(* IEC 61131-3 sources: kns-port-domestic/upstream/kns-pump-station/src/GVLs/Generated, 7 files *)

(* ---- GVL_CfgProject.gvl.st ---- *)
// AUTO-GENERATED by iolistgen 0.2.0 — не редактировать; источник: 03_io_list.csv
// SHA-256 перечня 06336d13c4b2; генератор st-codesys
// Назначение: уставки проекта — Cfg устройств из перечня сигналов, те же инициализаторы, что у GVL_Persist.
// PRG_ApplyProjectCfg копирует их в GVL_Persist (контракт plc-process-lib 18.3, правило 2).
{attribute 'qualified_only'}
VAR_GLOBAL CONSTANT
    // --- dev_no 11: P101 — Насос Н1 (MotorVfd) ---
    // lint:allow STL007 структура-константа: имя как у GVL_Persist.stP101Cfg (контракт 18.3, правило 2)
    stP101Cfg : PL.ST_MotorCfg := (
        tFbStart := T#10S,
        tFbStop := T#15S,
        tMinStop := T#30S,
        uiMaxStartsPerHour := 10,
        stVfd := (
            rSpeedMin_pct := 60.0,
            rRampUp_pctps := 5.0,
            rRampDown_pctps := 5.0,
            xFbFromComm := FALSE,
            xCommLossIsFault := FALSE
        ),
        udiAlarmIdBase := 110
    );
    // --- dev_no 12: P102 — Насос Н2 (MotorVfd) ---
    // lint:allow STL007 структура-константа: имя как у GVL_Persist.stP102Cfg (контракт 18.3, правило 2)
    stP102Cfg : PL.ST_MotorCfg := (
        tFbStart := T#10S,
        tFbStop := T#15S,
        tMinStop := T#30S,
        uiMaxStartsPerHour := 10,
        stVfd := (
            rSpeedMin_pct := 60.0,
            rRampUp_pctps := 5.0,
            rRampDown_pctps := 5.0,
            xFbFromComm := FALSE,
            xCommLossIsFault := FALSE
        ),
        udiAlarmIdBase := 120
    );
    // --- dev_no 13: P103 — Насос Н3 (MotorVfd) ---
    // lint:allow STL007 структура-константа: имя как у GVL_Persist.stP103Cfg (контракт 18.3, правило 2)
    stP103Cfg : PL.ST_MotorCfg := (
        tFbStart := T#10S,
        tFbStop := T#15S,
        tMinStop := T#30S,
        uiMaxStartsPerHour := 10,
        stVfd := (
            rSpeedMin_pct := 60.0,
            rRampUp_pctps := 5.0,
            rRampDown_pctps := 5.0,
            xFbFromComm := FALSE,
            xCommLossIsFault := FALSE
        ),
        udiAlarmIdBase := 130
    );
    // --- dev_no 14: V1 — Вытяжной вентилятор В1 павильона (Motor) ---
    // lint:allow STL007 структура-константа: имя как у GVL_Persist.stV1Cfg (контракт 18.3, правило 2)
    stV1Cfg : PL.ST_MotorCfg := (
        tMinStop := T#10S,
        udiAlarmIdBase := 140,
        astAlarm := [
            (ePriority := PL.E_AlarmPriority.Low),  // 0 FailToStart
            (ePriority := PL.E_AlarmPriority.Low),  // 1 FeedbackLost
            (ePriority := PL.E_AlarmPriority.High),  // 2 FailToStop
            (ePriority := PL.E_AlarmPriority.High),  // 3 UncommandedRun
            (ePriority := PL.E_AlarmPriority.Low),  // 4 ExtFault
            (ePriority := PL.E_AlarmPriority.None),  // 5 InterlockTrip
            (ePriority := PL.E_AlarmPriority.Medium),  // 6 CommLoss
            (ePriority := PL.E_AlarmPriority.Low)  // 7 SpeedDeviation
        ]
    );
    // --- dev_no 101: LT101 — Уровень в приёмном резервуаре (AnalogInput) ---
    // lint:allow STL007 структура-константа: имя как у GVL_Persist.stLT101Cfg (контракт 18.3, правило 2)
    stLT101Cfg : PL.ST_AnalogInputCfg := (
        rRangeHi_eu := 5.0,
        tFilter := T#2S,
        astLimit := [
            (xEnable := TRUE, rSetpoint_eu := 4.0, rHyst_eu := 0.05, tOnDelay := T#3S),  // 0 HH
            (xEnable := TRUE, rSetpoint_eu := 3.5, rHyst_eu := 0.05, tOnDelay := T#3S),  // 1 H
            (xEnable := TRUE, rSetpoint_eu := 0.8, rHyst_eu := 0.05, tOnDelay := T#3S),  // 2 L
            (xEnable := TRUE, rSetpoint_eu := 0.5, rHyst_eu := 0.05, tOnDelay := T#3S)  // 3 LL
        ],
        udiAlarmIdBase := 1010,
        astAlarm := [
            (ePriority := PL.E_AlarmPriority.High),  // 0 HH
            (ePriority := PL.E_AlarmPriority.Medium),  // 1 H
            (ePriority := PL.E_AlarmPriority.Medium),  // 2 L
            (ePriority := PL.E_AlarmPriority.High),  // 3 LL
            (ePriority := PL.E_AlarmPriority.Medium),  // 4 Failure
            (ePriority := PL.E_AlarmPriority.Low),  // 5 OutOfRange
            (ePriority := PL.E_AlarmPriority.None),  // 6 (резерв)
            (ePriority := PL.E_AlarmPriority.None)  // 7 (резерв)
        ]
    );
    // --- dev_no 102: LS102 — Поплавок «аварийно высокий уровень» (H, 4,2 м) (DigitalInput) ---
    // lint:allow STL007 структура-константа: имя как у GVL_Persist.stLS102Cfg (контракт 18.3, правило 2)
    stLS102Cfg : PL.ST_DigitalInputCfg := (
        xInvert := TRUE,
        tOnDelay := T#2S,
        udiAlarmIdBase := 1020,
        astAlarm := [
            (ePriority := PL.E_AlarmPriority.High),  // 0 State
            (ePriority := PL.E_AlarmPriority.Medium),  // 1 Failure
            (ePriority := PL.E_AlarmPriority.None),  // 2 (резерв)
            (ePriority := PL.E_AlarmPriority.None),  // 3 (резерв)
            (ePriority := PL.E_AlarmPriority.None),  // 4 (резерв)
            (ePriority := PL.E_AlarmPriority.None),  // 5 (резерв)
            (ePriority := PL.E_AlarmPriority.None),  // 6 (резерв)
            (ePriority := PL.E_AlarmPriority.None)  // 7 (резерв)
        ]
    );
    // --- dev_no 103: LS103 — Поплавок «сухой ход» (L, 0,4 м) (DigitalInput) ---
    // lint:allow STL007 структура-константа: имя как у GVL_Persist.stLS103Cfg (контракт 18.3, правило 2)
    stLS103Cfg : PL.ST_DigitalInputCfg := (
        xInvert := TRUE,
        tOnDelay := T#1S,
        eFailValue := PL.E_DiFailValue.ForceTrue,
        udiAlarmIdBase := 1030,
        astAlarm := [
            (ePriority := PL.E_AlarmPriority.High),  // 0 State
            (ePriority := PL.E_AlarmPriority.Medium),  // 1 Failure
            (ePriority := PL.E_AlarmPriority.None),  // 2 (резерв)
            (ePriority := PL.E_AlarmPriority.None),  // 3 (резерв)
            (ePriority := PL.E_AlarmPriority.None),  // 4 (резерв)
            (ePriority := PL.E_AlarmPriority.None),  // 5 (резерв)
            (ePriority := PL.E_AlarmPriority.None),  // 6 (резерв)
            (ePriority := PL.E_AlarmPriority.None)  // 7 (резерв)
        ]
    );
    // --- dev_no 111: IT111 — Насос Н1: ток двигателя (измеряет ПЧ) (AnalogInput) ---
    // lint:allow STL007 структура-константа: имя как у GVL_Persist.stIT111Cfg (контракт 18.3, правило 2)
    stIT111Cfg : PL.ST_AnalogInputCfg := (
        eInput := PL.E_AiInputType.Raw,
        rRangeHi_eu := 60.0,
        rRawHi_cnt := 600.0,
        tFilter := T#1S,
        astLimit := [
            (xEnable := TRUE, rSetpoint_eu := 34.0, tOnDelay := T#10S),  // 0 HH
            (xEnable := TRUE, rSetpoint_eu := 31.0, tOnDelay := T#10S),  // 1 H
            (xEnable := FALSE),  // 2 L
            (xEnable := FALSE)  // 3 LL
        ],
        udiAlarmIdBase := 1110,
        astAlarm := [
            (ePriority := PL.E_AlarmPriority.Medium),  // 0 HH
            (ePriority := PL.E_AlarmPriority.Low),  // 1 H
            (ePriority := PL.E_AlarmPriority.Low),  // 2 L
            (ePriority := PL.E_AlarmPriority.Medium),  // 3 LL
            (ePriority := PL.E_AlarmPriority.Medium),  // 4 Failure
            (ePriority := PL.E_AlarmPriority.Low),  // 5 OutOfRange
            (ePriority := PL.E_AlarmPriority.None),  // 6 (резерв)
            (ePriority := PL.E_AlarmPriority.None)  // 7 (резерв)
        ]
    );
    // --- dev_no 112: TS112 — Насос Н1: перегрев обмотки (термовыключатели, реле защиты насоса) (DigitalInput) ---
    // lint:allow STL007 структура-константа: имя как у GVL_Persist.stTS112Cfg (контракт 18.3, правило 2)
    stTS112Cfg : PL.ST_DigitalInputCfg := (
        xInvert := TRUE,
        udiAlarmIdBase := 1120,
        astAlarm := [
            (ePriority := PL.E_AlarmPriority.High),  // 0 State
            (ePriority := PL.E_AlarmPriority.Medium),  // 1 Failure
            (ePriority := PL.E_AlarmPriority.None),  // 2 (резерв)
            (ePriority := PL.E_AlarmPriority.None),  // 3 (резерв)
            (ePriority := PL.E_AlarmPriority.None),  // 4 (резерв)
            (ePriority := PL.E_AlarmPriority.None),  // 5 (резерв)
            (ePriority := PL.E_AlarmPriority.None),  // 6 (резерв)
            (ePriority := PL.E_AlarmPriority.None)  // 7 (резерв)
        ]
    );
    // --- dev_no 113: MS113 — Насос Н1: протечка в камеру статора (датчик влажности, реле защиты на… (DigitalInput) ---
    // lint:allow STL007 структура-константа: имя как у GVL_Persist.stMS113Cfg (контракт 18.3, правило 2)
    stMS113Cfg : PL.ST_DigitalInputCfg := (
        tOnDelay := T#10S,
        udiAlarmIdBase := 1130,
        astAlarm := [
            (ePriority := PL.E_AlarmPriority.Medium),  // 0 State
            (ePriority := PL.E_AlarmPriority.Medium),  // 1 Failure
            (ePriority := PL.E_AlarmPriority.None),  // 2 (резерв)
            (ePriority := PL.E_AlarmPriority.None),  // 3 (резерв)
            (ePriority := PL.E_AlarmPriority.None),  // 4 (резерв)
            (ePriority := PL.E_AlarmPriority.None),  // 5 (резерв)
            (ePriority := PL.E_AlarmPriority.None),  // 6 (резерв)
            (ePriority := PL.E_AlarmPriority.None)  // 7 (резерв)
        ]
    );
    // --- dev_no 121: IT121 — Насос Н2: ток двигателя (измеряет ПЧ) (AnalogInput) ---
    // lint:allow STL007 структура-константа: имя как у GVL_Persist.stIT121Cfg (контракт 18.3, правило 2)
    stIT121Cfg : PL.ST_AnalogInputCfg := (
        eInput := PL.E_AiInputType.Raw,
        rRangeHi_eu := 60.0,
        rRawHi_cnt := 600.0,
        tFilter := T#1S,
        astLimit := [
            (xEnable := TRUE, rSetpoint_eu := 34.0, tOnDelay := T#10S),  // 0 HH
            (xEnable := TRUE, rSetpoint_eu := 31.0, tOnDelay := T#10S),  // 1 H
            (xEnable := FALSE),  // 2 L
            (xEnable := FALSE)  // 3 LL
        ],
        udiAlarmIdBase := 1210,
        astAlarm := [
            (ePriority := PL.E_AlarmPriority.Medium),  // 0 HH
            (ePriority := PL.E_AlarmPriority.Low),  // 1 H
            (ePriority := PL.E_AlarmPriority.Low),  // 2 L
            (ePriority := PL.E_AlarmPriority.Medium),  // 3 LL
            (ePriority := PL.E_AlarmPriority.Medium),  // 4 Failure
            (ePriority := PL.E_AlarmPriority.Low),  // 5 OutOfRange
            (ePriority := PL.E_AlarmPriority.None),  // 6 (резерв)
            (ePriority := PL.E_AlarmPriority.None)  // 7 (резерв)
        ]
    );
    // --- dev_no 122: TS122 — Насос Н2: перегрев обмотки (термовыключатели, реле защиты насоса) (DigitalInput) ---
    // lint:allow STL007 структура-константа: имя как у GVL_Persist.stTS122Cfg (контракт 18.3, правило 2)
    stTS122Cfg : PL.ST_DigitalInputCfg := (
        xInvert := TRUE,
        udiAlarmIdBase := 1220,
        astAlarm := [
            (ePriority := PL.E_AlarmPriority.High),  // 0 State
            (ePriority := PL.E_AlarmPriority.Medium),  // 1 Failure
            (ePriority := PL.E_AlarmPriority.None),  // 2 (резерв)
            (ePriority := PL.E_AlarmPriority.None),  // 3 (резерв)
            (ePriority := PL.E_AlarmPriority.None),  // 4 (резерв)
            (ePriority := PL.E_AlarmPriority.None),  // 5 (резерв)
            (ePriority := PL.E_AlarmPriority.None),  // 6 (резерв)
            (ePriority := PL.E_AlarmPriority.None)  // 7 (резерв)
        ]
    );
    // --- dev_no 123: MS123 — Насос Н2: протечка в камеру статора (датчик влажности, реле защиты на… (DigitalInput) ---
    // lint:allow STL007 структура-константа: имя как у GVL_Persist.stMS123Cfg (контракт 18.3, правило 2)
    stMS123Cfg : PL.ST_DigitalInputCfg := (
        tOnDelay := T#10S,
        udiAlarmIdBase := 1230,
        astAlarm := [
            (ePriority := PL.E_AlarmPriority.Medium),  // 0 State
            (ePriority := PL.E_AlarmPriority.Medium),  // 1 Failure
            (ePriority := PL.E_AlarmPriority.None),  // 2 (резерв)
            (ePriority := PL.E_AlarmPriority.None),  // 3 (резерв)
            (ePriority := PL.E_AlarmPriority.None),  // 4 (резерв)
            (ePriority := PL.E_AlarmPriority.None),  // 5 (резерв)
            (ePriority := PL.E_AlarmPriority.None),  // 6 (резерв)
            (ePriority := PL.E_AlarmPriority.None)  // 7 (резерв)
        ]
    );
    // --- dev_no 131: IT131 — Насос Н3: ток двигателя (измеряет ПЧ) (AnalogInput) ---
    // lint:allow STL007 структура-константа: имя как у GVL_Persist.stIT131Cfg (контракт 18.3, правило 2)
    stIT131Cfg : PL.ST_AnalogInputCfg := (
        eInput := PL.E_AiInputType.Raw,
        rRangeHi_eu := 60.0,
        rRawHi_cnt := 600.0,
        tFilter := T#1S,
        astLimit := [
            (xEnable := TRUE, rSetpoint_eu := 34.0, tOnDelay := T#10S),  // 0 HH
            (xEnable := TRUE, rSetpoint_eu := 31.0, tOnDelay := T#10S),  // 1 H
            (xEnable := FALSE),  // 2 L
            (xEnable := FALSE)  // 3 LL
        ],
        udiAlarmIdBase := 1310,
        astAlarm := [
            (ePriority := PL.E_AlarmPriority.Medium),  // 0 HH
            (ePriority := PL.E_AlarmPriority.Low),  // 1 H
            (ePriority := PL.E_AlarmPriority.Low),  // 2 L
            (ePriority := PL.E_AlarmPriority.Medium),  // 3 LL
            (ePriority := PL.E_AlarmPriority.Medium),  // 4 Failure
            (ePriority := PL.E_AlarmPriority.Low),  // 5 OutOfRange
            (ePriority := PL.E_AlarmPriority.None),  // 6 (резерв)
            (ePriority := PL.E_AlarmPriority.None)  // 7 (резерв)
        ]
    );
    // --- dev_no 132: TS132 — Насос Н3: перегрев обмотки (термовыключатели, реле защиты насоса) (DigitalInput) ---
    // lint:allow STL007 структура-константа: имя как у GVL_Persist.stTS132Cfg (контракт 18.3, правило 2)
    stTS132Cfg : PL.ST_DigitalInputCfg := (
        xInvert := TRUE,
        udiAlarmIdBase := 1320,
        astAlarm := [
            (ePriority := PL.E_AlarmPriority.High),  // 0 State
            (ePriority := PL.E_AlarmPriority.Medium),  // 1 Failure
            (ePriority := PL.E_AlarmPriority.None),  // 2 (резерв)
            (ePriority := PL.E_AlarmPriority.None),  // 3 (резерв)
            (ePriority := PL.E_AlarmPriority.None),  // 4 (резерв)
            (ePriority := PL.E_AlarmPriority.None),  // 5 (резерв)
            (ePriority := PL.E_AlarmPriority.None),  // 6 (резерв)
            (ePriority := PL.E_AlarmPriority.None)  // 7 (резерв)
        ]
    );
    // --- dev_no 133: MS133 — Насос Н3: протечка в камеру статора (датчик влажности, реле защиты на… (DigitalInput) ---
    // lint:allow STL007 структура-константа: имя как у GVL_Persist.stMS133Cfg (контракт 18.3, правило 2)
    stMS133Cfg : PL.ST_DigitalInputCfg := (
        tOnDelay := T#10S,
        udiAlarmIdBase := 1330,
        astAlarm := [
            (ePriority := PL.E_AlarmPriority.Medium),  // 0 State
            (ePriority := PL.E_AlarmPriority.Medium),  // 1 Failure
            (ePriority := PL.E_AlarmPriority.None),  // 2 (резерв)
            (ePriority := PL.E_AlarmPriority.None),  // 3 (резерв)
            (ePriority := PL.E_AlarmPriority.None),  // 4 (резерв)
            (ePriority := PL.E_AlarmPriority.None),  // 5 (резерв)
            (ePriority := PL.E_AlarmPriority.None),  // 6 (резерв)
            (ePriority := PL.E_AlarmPriority.None)  // 7 (резерв)
        ]
    );
    // --- dev_no 201: PT201 — Давление в напорном коллекторе (AnalogInput) ---
    // lint:allow STL007 структура-константа: имя как у GVL_Persist.stPT201Cfg (контракт 18.3, правило 2)
    stPT201Cfg : PL.ST_AnalogInputCfg := (
        rRangeHi_eu := 10.0,
        tFilter := T#1S,
        astLimit := [
            (xEnable := TRUE, rSetpoint_eu := 5.0, tOnDelay := T#5S),  // 0 HH
            (xEnable := TRUE, rSetpoint_eu := 4.0, tOnDelay := T#5S),  // 1 H
            (xEnable := TRUE, rSetpoint_eu := 1.0, rHyst_eu := 0.1, tOnDelay := T#5S),  // 2 L
            (xEnable := TRUE, rSetpoint_eu := 0.5, rHyst_eu := 0.1, tOnDelay := T#5S)  // 3 LL
        ],
        udiAlarmIdBase := 2010,
        astAlarm := [
            (ePriority := PL.E_AlarmPriority.High),  // 0 HH
            (ePriority := PL.E_AlarmPriority.Medium),  // 1 H
            (ePriority := PL.E_AlarmPriority.Medium),  // 2 L
            (ePriority := PL.E_AlarmPriority.High),  // 3 LL
            (ePriority := PL.E_AlarmPriority.Medium),  // 4 Failure
            (ePriority := PL.E_AlarmPriority.Low),  // 5 OutOfRange
            (ePriority := PL.E_AlarmPriority.None),  // 6 (резерв)
            (ePriority := PL.E_AlarmPriority.None)  // 7 (резерв)
        ]
    );
    // --- dev_no 202: FT202 — Расход в напорном коллекторе (AnalogInput) ---
    // lint:allow STL007 структура-константа: имя как у GVL_Persist.stFT202Cfg (контракт 18.3, правило 2)
    stFT202Cfg : PL.ST_AnalogInputCfg := (
        rRangeHi_eu := 500.0,
        rLowCut_pct := 1.0,
        tFilter := T#3S,
        astLimit := [
            (xEnable := FALSE),  // 0 HH
            (xEnable := FALSE),  // 1 H
            (xEnable := TRUE, rSetpoint_eu := 30.0, rHyst_eu := 5.0, tOnDelay := T#30S),  // 2 L
            (xEnable := FALSE)  // 3 LL
        ],
        udiAlarmIdBase := 2020,
        astAlarm := [
            (ePriority := PL.E_AlarmPriority.High),  // 0 HH
            (ePriority := PL.E_AlarmPriority.Low),  // 1 H
            (ePriority := PL.E_AlarmPriority.Medium),  // 2 L
            (ePriority := PL.E_AlarmPriority.High),  // 3 LL
            (ePriority := PL.E_AlarmPriority.Medium),  // 4 Failure
            (ePriority := PL.E_AlarmPriority.Low),  // 5 OutOfRange
            (ePriority := PL.E_AlarmPriority.None),  // 6 (резерв)
            (ePriority := PL.E_AlarmPriority.None)  // 7 (резерв)
        ]
    );
    // --- dev_no 203: LS203 — Затопление камеры задвижек (DigitalInput) ---
    // lint:allow STL007 структура-константа: имя как у GVL_Persist.stLS203Cfg (контракт 18.3, правило 2)
    stLS203Cfg : PL.ST_DigitalInputCfg := (
        tOnDelay := T#5S,
        udiAlarmIdBase := 2030,
        astAlarm := [
            (ePriority := PL.E_AlarmPriority.Medium),  // 0 State
            (ePriority := PL.E_AlarmPriority.Medium),  // 1 Failure
            (ePriority := PL.E_AlarmPriority.None),  // 2 (резерв)
            (ePriority := PL.E_AlarmPriority.None),  // 3 (резерв)
            (ePriority := PL.E_AlarmPriority.None),  // 4 (резерв)
            (ePriority := PL.E_AlarmPriority.None),  // 5 (резерв)
            (ePriority := PL.E_AlarmPriority.None),  // 6 (резерв)
            (ePriority := PL.E_AlarmPriority.None)  // 7 (резерв)
        ]
    );
    // --- dev_no 301: ES301 — Напряжение на вводе в норме (реле контроля фаз) (DigitalInput) ---
    // lint:allow STL007 структура-константа: имя как у GVL_Persist.stES301Cfg (контракт 18.3, правило 2)
    stES301Cfg : PL.ST_DigitalInputCfg := (
        tOnDelay := T#3S,
        xAlarmOnTrue := FALSE,
        udiAlarmIdBase := 3010,
        astAlarm := [
            (ePriority := PL.E_AlarmPriority.High),  // 0 State
            (ePriority := PL.E_AlarmPriority.Medium),  // 1 Failure
            (ePriority := PL.E_AlarmPriority.None),  // 2 (резерв)
            (ePriority := PL.E_AlarmPriority.None),  // 3 (резерв)
            (ePriority := PL.E_AlarmPriority.None),  // 4 (резерв)
            (ePriority := PL.E_AlarmPriority.None),  // 5 (резерв)
            (ePriority := PL.E_AlarmPriority.None),  // 6 (резерв)
            (ePriority := PL.E_AlarmPriority.None)  // 7 (резерв)
        ]
    );
    // --- dev_no 302: YS302 — ИБП шкафа управления: работа от батарей (DigitalInput) ---
    // lint:allow STL007 структура-константа: имя как у GVL_Persist.stYS302Cfg (контракт 18.3, правило 2)
    stYS302Cfg : PL.ST_DigitalInputCfg := (
        tOnDelay := T#5S,
        udiAlarmIdBase := 3020,
        astAlarm := [
            (ePriority := PL.E_AlarmPriority.Medium),  // 0 State
            (ePriority := PL.E_AlarmPriority.Medium),  // 1 Failure
            (ePriority := PL.E_AlarmPriority.None),  // 2 (резерв)
            (ePriority := PL.E_AlarmPriority.None),  // 3 (резерв)
            (ePriority := PL.E_AlarmPriority.None),  // 4 (резерв)
            (ePriority := PL.E_AlarmPriority.None),  // 5 (резерв)
            (ePriority := PL.E_AlarmPriority.None),  // 6 (резерв)
            (ePriority := PL.E_AlarmPriority.None)  // 7 (резерв)
        ]
    );
    // --- dev_no 303: YS303 — ИБП шкафа управления: неисправность или разряд батарей (DigitalInput) ---
    // lint:allow STL007 структура-константа: имя как у GVL_Persist.stYS303Cfg (контракт 18.3, правило 2)
    stYS303Cfg : PL.ST_DigitalInputCfg := (
        tOnDelay := T#5S,
        udiAlarmIdBase := 3030,
        astAlarm := [
            (ePriority := PL.E_AlarmPriority.Medium),  // 0 State
            (ePriority := PL.E_AlarmPriority.Medium),  // 1 Failure
            (ePriority := PL.E_AlarmPriority.None),  // 2 (резерв)
            (ePriority := PL.E_AlarmPriority.None),  // 3 (резерв)
            (ePriority := PL.E_AlarmPriority.None),  // 4 (резерв)
            (ePriority := PL.E_AlarmPriority.None),  // 5 (резерв)
            (ePriority := PL.E_AlarmPriority.None),  // 6 (резерв)
            (ePriority := PL.E_AlarmPriority.None)  // 7 (резерв)
        ]
    );
    // --- dev_no 401: AT401 — Концентрация сероводорода H₂S в павильоне (AnalogInput) ---
    // lint:allow STL007 структура-константа: имя как у GVL_Persist.stAT401Cfg (контракт 18.3, правило 2)
    stAT401Cfg : PL.ST_AnalogInputCfg := (
        rRangeHi_eu := 40.0,
        astLimit := [
            (xEnable := TRUE, rSetpoint_eu := 10.0, rHyst_eu := 0.5, tOnDelay := T#5S),  // 0 HH
            (xEnable := TRUE, rSetpoint_eu := 5.0, rHyst_eu := 0.5, tOnDelay := T#5S),  // 1 H
            (xEnable := FALSE),  // 2 L
            (xEnable := FALSE)  // 3 LL
        ],
        udiAlarmIdBase := 4010,
        astAlarm := [
            (ePriority := PL.E_AlarmPriority.High),  // 0 HH
            (ePriority := PL.E_AlarmPriority.Medium),  // 1 H
            (ePriority := PL.E_AlarmPriority.Medium),  // 2 L
            (ePriority := PL.E_AlarmPriority.High),  // 3 LL
            (ePriority := PL.E_AlarmPriority.Medium),  // 4 Failure
            (ePriority := PL.E_AlarmPriority.Low),  // 5 OutOfRange
            (ePriority := PL.E_AlarmPriority.None),  // 6 (резерв)
            (ePriority := PL.E_AlarmPriority.None)  // 7 (резерв)
        ]
    );
    // --- dev_no 402: AT402 — Концентрация метана CH₄ в павильоне (AnalogInput) ---
    // lint:allow STL007 структура-константа: имя как у GVL_Persist.stAT402Cfg (контракт 18.3, правило 2)
    stAT402Cfg : PL.ST_AnalogInputCfg := (
        astLimit := [
            (xEnable := TRUE, rSetpoint_eu := 20.0, rHyst_eu := 1.0, tOnDelay := T#5S),  // 0 HH
            (xEnable := TRUE, rSetpoint_eu := 10.0, rHyst_eu := 1.0, tOnDelay := T#5S),  // 1 H
            (xEnable := FALSE),  // 2 L
            (xEnable := FALSE)  // 3 LL
        ],
        udiAlarmIdBase := 4020,
        astAlarm := [
            (ePriority := PL.E_AlarmPriority.High),  // 0 HH
            (ePriority := PL.E_AlarmPriority.Medium),  // 1 H
            (ePriority := PL.E_AlarmPriority.Medium),  // 2 L
            (ePriority := PL.E_AlarmPriority.High),  // 3 LL
            (ePriority := PL.E_AlarmPriority.Medium),  // 4 Failure
            (ePriority := PL.E_AlarmPriority.Low),  // 5 OutOfRange
            (ePriority := PL.E_AlarmPriority.None),  // 6 (резерв)
            (ePriority := PL.E_AlarmPriority.None)  // 7 (резерв)
        ]
    );
    // --- dev_no 403: TT403 — Температура воздуха в павильоне (AnalogInput) ---
    // lint:allow STL007 структура-константа: имя как у GVL_Persist.stTT403Cfg (контракт 18.3, правило 2)
    stTT403Cfg : PL.ST_AnalogInputCfg := (
        eInput := PL.E_AiInputType.Eng,
        rRangeLo_eu := -40.0,
        rRangeHi_eu := 60.0,
        astLimit := [
            (xEnable := FALSE),  // 0 HH
            (xEnable := TRUE, rSetpoint_eu := 35.0, rHyst_eu := 1.0, tOnDelay := T#1M),  // 1 H
            (xEnable := TRUE, rSetpoint_eu := 5.0, rHyst_eu := 1.0, tOnDelay := T#1M),  // 2 L
            (xEnable := FALSE)  // 3 LL
        ],
        udiAlarmIdBase := 4030,
        astAlarm := [
            (ePriority := PL.E_AlarmPriority.Low),  // 0 HH
            (ePriority := PL.E_AlarmPriority.Low),  // 1 H
            (ePriority := PL.E_AlarmPriority.Low),  // 2 L
            (ePriority := PL.E_AlarmPriority.Low),  // 3 LL
            (ePriority := PL.E_AlarmPriority.Medium),  // 4 Failure
            (ePriority := PL.E_AlarmPriority.Low),  // 5 OutOfRange
            (ePriority := PL.E_AlarmPriority.None),  // 6 (резерв)
            (ePriority := PL.E_AlarmPriority.None)  // 7 (резерв)
        ]
    );
    // --- dev_no 404: ZS404 — Дверь павильона открыта (DigitalInput) ---
    // lint:allow STL007 структура-константа: имя как у GVL_Persist.stZS404Cfg (контракт 18.3, правило 2)
    stZS404Cfg : PL.ST_DigitalInputCfg := (
        tOnDelay := T#2S,
        udiAlarmIdBase := 4040,
        astAlarm := [
            (ePriority := PL.E_AlarmPriority.Low),  // 0 State
            (ePriority := PL.E_AlarmPriority.Medium),  // 1 Failure
            (ePriority := PL.E_AlarmPriority.None),  // 2 (резерв)
            (ePriority := PL.E_AlarmPriority.None),  // 3 (резерв)
            (ePriority := PL.E_AlarmPriority.None),  // 4 (резерв)
            (ePriority := PL.E_AlarmPriority.None),  // 5 (резерв)
            (ePriority := PL.E_AlarmPriority.None),  // 6 (резерв)
            (ePriority := PL.E_AlarmPriority.None)  // 7 (резерв)
        ]
    );
    // --- dev_no 405: YS405 — Пожар (сигнал прибора пожарной сигнализации) (DigitalInput) ---
    // lint:allow STL007 структура-константа: имя как у GVL_Persist.stYS405Cfg (контракт 18.3, правило 2)
    stYS405Cfg : PL.ST_DigitalInputCfg := (
        udiAlarmIdBase := 4050,
        astAlarm := [
            (ePriority := PL.E_AlarmPriority.High),  // 0 State
            (ePriority := PL.E_AlarmPriority.Medium),  // 1 Failure
            (ePriority := PL.E_AlarmPriority.None),  // 2 (резерв)
            (ePriority := PL.E_AlarmPriority.None),  // 3 (резерв)
            (ePriority := PL.E_AlarmPriority.None),  // 4 (резерв)
            (ePriority := PL.E_AlarmPriority.None),  // 5 (резерв)
            (ePriority := PL.E_AlarmPriority.None),  // 6 (резерв)
            (ePriority := PL.E_AlarmPriority.None)  // 7 (резерв)
        ]
    );
    // --- dev_no 501: HS501 — Кнопка «Сброс аварий» на двери шкафа управления (DigitalInput) ---
    // lint:allow STL007 структура-константа: имя как у GVL_Persist.stHS501Cfg (контракт 18.3, правило 2)
    stHS501Cfg : PL.ST_DigitalInputCfg := (udiAlarmIdBase := 5010);
    // --- dev_no 502: HS502 — Кнопка «Отключить звук» на двери шкафа управления (DigitalInput) ---
    // lint:allow STL007 структура-константа: имя как у GVL_Persist.stHS502Cfg (контракт 18.3, правило 2)
    stHS502Cfg : PL.ST_DigitalInputCfg := (udiAlarmIdBase := 5020);
END_VAR

(* ---- GVL_DeviceList.gvl.st ---- *)
// AUTO-GENERATED by tools_project/generate.py — не редактировать; источник: docs/03_io_list.csv
// Назначение: список устройств перечня для общего сброса и квитирования, сводки тревог, аудита режимов
//             и кодов тревог в CSV журнала (решение D-11): теги, dev_no и типы по возрастанию dev_no,
//             позиция устройства в списке (IDX_<TAG>) и интерфейсы aitfDevice, которые присваивает
//             PRG_DeviceList каждый цикл (ссылки переживают онлайн-изменение).
{attribute 'qualified_only'}
VAR_GLOBAL CONSTANT
    DEVICE_COUNT : UINT := 29;  // устройств в перечне сигналов
    IDX_P101 : UINT := 1;  // 11 · Насос Н1
    IDX_P102 : UINT := 2;  // 12 · Насос Н2
    IDX_P103 : UINT := 3;  // 13 · Насос Н3
    IDX_V1 : UINT := 4;  // 14 · Вытяжной вентилятор В1 павильона
    IDX_LT101 : UINT := 5;  // 101 · Уровень в приёмном резервуаре
    IDX_LS102 : UINT := 6;  // 102 · Поплавок «аварийно высокий уровень» (H, 4,2 м)
    IDX_LS103 : UINT := 7;  // 103 · Поплавок «сухой ход» (L, 0,4 м)
    IDX_IT111 : UINT := 8;  // 111 · Насос Н1: ток двигателя (измеряет ПЧ)
    IDX_TS112 : UINT := 9;  // 112 · Насос Н1: перегрев обмотки (термовыключатели, реле защиты насоса)
    IDX_MS113 : UINT := 10;  // 113 · Насос Н1: протечка в камеру статора (датчик влажности, реле защиты насоса)
    IDX_IT121 : UINT := 11;  // 121 · Насос Н2: ток двигателя (измеряет ПЧ)
    IDX_TS122 : UINT := 12;  // 122 · Насос Н2: перегрев обмотки (термовыключатели, реле защиты насоса)
    IDX_MS123 : UINT := 13;  // 123 · Насос Н2: протечка в камеру статора (датчик влажности, реле защиты насоса)
    IDX_IT131 : UINT := 14;  // 131 · Насос Н3: ток двигателя (измеряет ПЧ)
    IDX_TS132 : UINT := 15;  // 132 · Насос Н3: перегрев обмотки (термовыключатели, реле защиты насоса)
    IDX_MS133 : UINT := 16;  // 133 · Насос Н3: протечка в камеру статора (датчик влажности, реле защиты насоса)
    IDX_PT201 : UINT := 17;  // 201 · Давление в напорном коллекторе
    IDX_FT202 : UINT := 18;  // 202 · Расход в напорном коллекторе
    IDX_LS203 : UINT := 19;  // 203 · Затопление камеры задвижек
    IDX_ES301 : UINT := 20;  // 301 · Напряжение на вводе в норме (реле контроля фаз)
    IDX_YS302 : UINT := 21;  // 302 · ИБП шкафа управления: работа от батарей
    IDX_YS303 : UINT := 22;  // 303 · ИБП шкафа управления: неисправность или разряд батарей
    IDX_AT401 : UINT := 23;  // 401 · Концентрация сероводорода H₂S в павильоне
    IDX_AT402 : UINT := 24;  // 402 · Концентрация метана CH₄ в павильоне
    IDX_TT403 : UINT := 25;  // 403 · Температура воздуха в павильоне
    IDX_ZS404 : UINT := 26;  // 404 · Дверь павильона открыта
    IDX_YS405 : UINT := 27;  // 405 · Пожар (сигнал прибора пожарной сигнализации)
    IDX_HS501 : UINT := 28;  // 501 · Кнопка «Сброс аварий» на двери шкафа управления
    IDX_HS502 : UINT := 29;  // 502 · Кнопка «Отключить звук» на двери шкафа управления
    // lint:allow STL007 имя как у переменной списка (DESIGN, раздел 4.5): массив-константа
    asTag : ARRAY[1..GVL_DeviceList.DEVICE_COUNT] OF STRING(GVL_Const.TAG_LEN) := ['P101', 'P102', 'P103', 'V1',
        'LT101', 'LS102', 'LS103', 'IT111', 'TS112', 'MS113', 'IT121', 'TS122', 'MS123', 'IT131', 'TS132', 'MS133',
        'PT201', 'FT202', 'LS203', 'ES301', 'YS302', 'YS303', 'AT401', 'AT402', 'TT403', 'ZS404', 'YS405', 'HS501',
        'HS502'];
    // lint:allow STL007 имя как у переменной списка (DESIGN, раздел 4.5): массив-константа
    auiDevNo : ARRAY[1..GVL_DeviceList.DEVICE_COUNT] OF UINT := [GVL_DevIdx.P101, GVL_DevIdx.P102, GVL_DevIdx.P103,
        GVL_DevIdx.V1, GVL_DevIdx.LT101, GVL_DevIdx.LS102, GVL_DevIdx.LS103, GVL_DevIdx.IT111, GVL_DevIdx.TS112,
        GVL_DevIdx.MS113, GVL_DevIdx.IT121, GVL_DevIdx.TS122, GVL_DevIdx.MS123, GVL_DevIdx.IT131, GVL_DevIdx.TS132,
        GVL_DevIdx.MS133, GVL_DevIdx.PT201, GVL_DevIdx.FT202, GVL_DevIdx.LS203, GVL_DevIdx.ES301, GVL_DevIdx.YS302,
        GVL_DevIdx.YS303, GVL_DevIdx.AT401, GVL_DevIdx.AT402, GVL_DevIdx.TT403, GVL_DevIdx.ZS404, GVL_DevIdx.YS405,
        GVL_DevIdx.HS501, GVL_DevIdx.HS502];
    // lint:allow STL007 имя как у переменной списка (DESIGN, раздел 4.5): массив-константа
    aeDevType : ARRAY[1..GVL_DeviceList.DEVICE_COUNT] OF PL.E_DeviceType := [PL.E_DeviceType.MotorVfd,
        PL.E_DeviceType.MotorVfd, PL.E_DeviceType.MotorVfd, PL.E_DeviceType.Motor, PL.E_DeviceType.AnalogInput,
        PL.E_DeviceType.DigitalInput, PL.E_DeviceType.DigitalInput, PL.E_DeviceType.AnalogInput,
        PL.E_DeviceType.DigitalInput, PL.E_DeviceType.DigitalInput, PL.E_DeviceType.AnalogInput,
        PL.E_DeviceType.DigitalInput, PL.E_DeviceType.DigitalInput, PL.E_DeviceType.AnalogInput,
        PL.E_DeviceType.DigitalInput, PL.E_DeviceType.DigitalInput, PL.E_DeviceType.AnalogInput,
        PL.E_DeviceType.AnalogInput, PL.E_DeviceType.DigitalInput, PL.E_DeviceType.DigitalInput,
        PL.E_DeviceType.DigitalInput, PL.E_DeviceType.DigitalInput, PL.E_DeviceType.AnalogInput,
        PL.E_DeviceType.AnalogInput, PL.E_DeviceType.AnalogInput, PL.E_DeviceType.DigitalInput,
        PL.E_DeviceType.DigitalInput, PL.E_DeviceType.DigitalInput, PL.E_DeviceType.DigitalInput];
END_VAR
VAR_GLOBAL
    aitfDevice : ARRAY[1..GVL_DeviceList.DEVICE_COUNT] OF PL.I_Device;  // присваивает PRG_DeviceList каждый цикл
END_VAR

(* ---- GVL_Devices.gvl.st ---- *)
// AUTO-GENERATED by iolistgen 0.2.0 — не редактировать; источник: 03_io_list.csv
// SHA-256 перечня 06336d13c4b2; генератор st-codesys
// Назначение: экземпляры устройств plc-process-lib (объявление без параметров, контракт 20). Логика станции пишет их
// входы автоматики и читает выходы; HMI и SCADA читают stSts.
{attribute 'qualified_only'}
VAR_GLOBAL
    fbP101 : PL.FB_MotorVfd;  // 11 · Насос Н1
    fbP102 : PL.FB_MotorVfd;  // 12 · Насос Н2
    fbP103 : PL.FB_MotorVfd;  // 13 · Насос Н3
    fbV1 : PL.FB_Motor;  // 14 · Вытяжной вентилятор В1 павильона
    fbLT101 : PL.FB_AnalogInput;  // 101 · Уровень в приёмном резервуаре
    fbLS102 : PL.FB_DigitalInput;  // 102 · Поплавок «аварийно высокий уровень» (H, 4,2 м)
    fbLS103 : PL.FB_DigitalInput;  // 103 · Поплавок «сухой ход» (L, 0,4 м)
    fbIT111 : PL.FB_AnalogInput;  // 111 · Насос Н1: ток двигателя (измеряет ПЧ)
    fbTS112 : PL.FB_DigitalInput;  // 112 · Насос Н1: перегрев обмотки (термовыключатели, реле защиты насоса)
    fbMS113 : PL.FB_DigitalInput;  // 113 · Насос Н1: протечка в камеру статора (датчик влажности, реле защиты насоса)
    fbIT121 : PL.FB_AnalogInput;  // 121 · Насос Н2: ток двигателя (измеряет ПЧ)
    fbTS122 : PL.FB_DigitalInput;  // 122 · Насос Н2: перегрев обмотки (термовыключатели, реле защиты насоса)
    fbMS123 : PL.FB_DigitalInput;  // 123 · Насос Н2: протечка в камеру статора (датчик влажности, реле защиты насоса)
    fbIT131 : PL.FB_AnalogInput;  // 131 · Насос Н3: ток двигателя (измеряет ПЧ)
    fbTS132 : PL.FB_DigitalInput;  // 132 · Насос Н3: перегрев обмотки (термовыключатели, реле защиты насоса)
    fbMS133 : PL.FB_DigitalInput;  // 133 · Насос Н3: протечка в камеру статора (датчик влажности, реле защиты насоса)
    fbPT201 : PL.FB_AnalogInput;  // 201 · Давление в напорном коллекторе
    fbFT202 : PL.FB_AnalogInput;  // 202 · Расход в напорном коллекторе
    fbLS203 : PL.FB_DigitalInput;  // 203 · Затопление камеры задвижек
    fbES301 : PL.FB_DigitalInput;  // 301 · Напряжение на вводе в норме (реле контроля фаз)
    fbYS302 : PL.FB_DigitalInput;  // 302 · ИБП шкафа управления: работа от батарей
    fbYS303 : PL.FB_DigitalInput;  // 303 · ИБП шкафа управления: неисправность или разряд батарей
    fbAT401 : PL.FB_AnalogInput;  // 401 · Концентрация сероводорода H₂S в павильоне
    fbAT402 : PL.FB_AnalogInput;  // 402 · Концентрация метана CH₄ в павильоне
    fbTT403 : PL.FB_AnalogInput;  // 403 · Температура воздуха в павильоне
    fbZS404 : PL.FB_DigitalInput;  // 404 · Дверь павильона открыта
    fbYS405 : PL.FB_DigitalInput;  // 405 · Пожар (сигнал прибора пожарной сигнализации)
    fbHS501 : PL.FB_DigitalInput;  // 501 · Кнопка «Сброс аварий» на двери шкафа управления
    fbHS502 : PL.FB_DigitalInput;  // 502 · Кнопка «Отключить звук» на двери шкафа управления
END_VAR

(* ---- GVL_DevIdx.gvl.st ---- *)
// AUTO-GENERATED by iolistgen 0.2.0 — не редактировать; источник: 03_io_list.csv
// SHA-256 перечня 06336d13c4b2; генератор st-codesys
// Назначение: номера устройств dev_no (контракт plc-process-lib 20.1): тревоги устройства — dev_no · 10 + слот; для
// SCADA и логики станции.
{attribute 'qualified_only'}
VAR_GLOBAL CONSTANT
    P101 : UINT := 11;  // MotorVfd · Насос Н1
    P102 : UINT := 12;  // MotorVfd · Насос Н2
    P103 : UINT := 13;  // MotorVfd · Насос Н3
    V1 : UINT := 14;  // Motor · Вытяжной вентилятор В1 павильона
    LT101 : UINT := 101;  // AnalogInput · Уровень в приёмном резервуаре
    LS102 : UINT := 102;  // DigitalInput · Поплавок «аварийно высокий уровень» (H, 4,2 м)
    LS103 : UINT := 103;  // DigitalInput · Поплавок «сухой ход» (L, 0,4 м)
    IT111 : UINT := 111;  // AnalogInput · Насос Н1: ток двигателя (измеряет ПЧ)
    TS112 : UINT := 112;  // DigitalInput · Насос Н1: перегрев обмотки (термовыключатели, реле защиты насоса)
    MS113 : UINT := 113;  // DigitalInput · Насос Н1: протечка в камеру статора (датчик влажности, реле защиты насоса)
    IT121 : UINT := 121;  // AnalogInput · Насос Н2: ток двигателя (измеряет ПЧ)
    TS122 : UINT := 122;  // DigitalInput · Насос Н2: перегрев обмотки (термовыключатели, реле защиты насоса)
    MS123 : UINT := 123;  // DigitalInput · Насос Н2: протечка в камеру статора (датчик влажности, реле защиты насоса)
    IT131 : UINT := 131;  // AnalogInput · Насос Н3: ток двигателя (измеряет ПЧ)
    TS132 : UINT := 132;  // DigitalInput · Насос Н3: перегрев обмотки (термовыключатели, реле защиты насоса)
    MS133 : UINT := 133;  // DigitalInput · Насос Н3: протечка в камеру статора (датчик влажности, реле защиты насоса)
    PT201 : UINT := 201;  // AnalogInput · Давление в напорном коллекторе
    FT202 : UINT := 202;  // AnalogInput · Расход в напорном коллекторе
    LS203 : UINT := 203;  // DigitalInput · Затопление камеры задвижек
    ES301 : UINT := 301;  // DigitalInput · Напряжение на вводе в норме (реле контроля фаз)
    YS302 : UINT := 302;  // DigitalInput · ИБП шкафа управления: работа от батарей
    YS303 : UINT := 303;  // DigitalInput · ИБП шкафа управления: неисправность или разряд батарей
    AT401 : UINT := 401;  // AnalogInput · Концентрация сероводорода H₂S в павильоне
    AT402 : UINT := 402;  // AnalogInput · Концентрация метана CH₄ в павильоне
    TT403 : UINT := 403;  // AnalogInput · Температура воздуха в павильоне
    ZS404 : UINT := 404;  // DigitalInput · Дверь павильона открыта
    YS405 : UINT := 405;  // DigitalInput · Пожар (сигнал прибора пожарной сигнализации)
    HS501 : UINT := 501;  // DigitalInput · Кнопка «Сброс аварий» на двери шкафа управления
    HS502 : UINT := 502;  // DigitalInput · Кнопка «Отключить звук» на двери шкафа управления
END_VAR

(* ---- GVL_Hmi.gvl.st ---- *)
// AUTO-GENERATED by iolistgen 0.2.0 — не редактировать; источник: 03_io_list.csv
// SHA-256 перечня 06336d13c4b2; генератор st-codesys
// Назначение: команды HMI и SCADA устройствам (ST_<Dev>Cmd, контракт plc-process-lib 1 и 2.1). WebVisu и OPC UA пишут
// сюда напрямую; команды по Modbus — только через адаптер приложения (импульс по фронту).
{attribute 'qualified_only'}
VAR_GLOBAL
    xApplyProjectCfg : BOOL;  // импульс: применить уставки проекта (PRG_ApplyProjectCfg); сбрасывает PRG_Devices
    stP101Cmd : PL.ST_MotorCmd;  // 11 · Насос Н1
    stP102Cmd : PL.ST_MotorCmd;  // 12 · Насос Н2
    stP103Cmd : PL.ST_MotorCmd;  // 13 · Насос Н3
    stV1Cmd : PL.ST_MotorCmd;  // 14 · Вытяжной вентилятор В1 павильона
    stLT101Cmd : PL.ST_AnalogInputCmd;  // 101 · Уровень в приёмном резервуаре
    stLS102Cmd : PL.ST_DigitalInputCmd;  // 102 · Поплавок «аварийно высокий уровень» (H, 4,2 м)
    stLS103Cmd : PL.ST_DigitalInputCmd;  // 103 · Поплавок «сухой ход» (L, 0,4 м)
    stIT111Cmd : PL.ST_AnalogInputCmd;  // 111 · Насос Н1: ток двигателя (измеряет ПЧ)
    stTS112Cmd : PL.ST_DigitalInputCmd;  // 112 · Насос Н1: перегрев обмотки (термовыключатели, реле защиты насоса)
    // 113 · Насос Н1: протечка в камеру статора (датчик влажности, реле защиты насоса)
    stMS113Cmd : PL.ST_DigitalInputCmd;
    stIT121Cmd : PL.ST_AnalogInputCmd;  // 121 · Насос Н2: ток двигателя (измеряет ПЧ)
    stTS122Cmd : PL.ST_DigitalInputCmd;  // 122 · Насос Н2: перегрев обмотки (термовыключатели, реле защиты насоса)
    // 123 · Насос Н2: протечка в камеру статора (датчик влажности, реле защиты насоса)
    stMS123Cmd : PL.ST_DigitalInputCmd;
    stIT131Cmd : PL.ST_AnalogInputCmd;  // 131 · Насос Н3: ток двигателя (измеряет ПЧ)
    stTS132Cmd : PL.ST_DigitalInputCmd;  // 132 · Насос Н3: перегрев обмотки (термовыключатели, реле защиты насоса)
    // 133 · Насос Н3: протечка в камеру статора (датчик влажности, реле защиты насоса)
    stMS133Cmd : PL.ST_DigitalInputCmd;
    stPT201Cmd : PL.ST_AnalogInputCmd;  // 201 · Давление в напорном коллекторе
    stFT202Cmd : PL.ST_AnalogInputCmd;  // 202 · Расход в напорном коллекторе
    stLS203Cmd : PL.ST_DigitalInputCmd;  // 203 · Затопление камеры задвижек
    stES301Cmd : PL.ST_DigitalInputCmd;  // 301 · Напряжение на вводе в норме (реле контроля фаз)
    stYS302Cmd : PL.ST_DigitalInputCmd;  // 302 · ИБП шкафа управления: работа от батарей
    stYS303Cmd : PL.ST_DigitalInputCmd;  // 303 · ИБП шкафа управления: неисправность или разряд батарей
    stAT401Cmd : PL.ST_AnalogInputCmd;  // 401 · Концентрация сероводорода H₂S в павильоне
    stAT402Cmd : PL.ST_AnalogInputCmd;  // 402 · Концентрация метана CH₄ в павильоне
    stTT403Cmd : PL.ST_AnalogInputCmd;  // 403 · Температура воздуха в павильоне
    stZS404Cmd : PL.ST_DigitalInputCmd;  // 404 · Дверь павильона открыта
    stYS405Cmd : PL.ST_DigitalInputCmd;  // 405 · Пожар (сигнал прибора пожарной сигнализации)
    stHS501Cmd : PL.ST_DigitalInputCmd;  // 501 · Кнопка «Сброс аварий» на двери шкафа управления
    stHS502Cmd : PL.ST_DigitalInputCmd;  // 502 · Кнопка «Отключить звук» на двери шкафа управления
END_VAR

(* ---- GVL_IO.gvl.st ---- *)
// AUTO-GENERATED by iolistgen 0.2.0 — не редактировать; источник: 03_io_list.csv
// SHA-256 перечня 06336d13c4b2; генератор st-codesys
// Назначение: переменные ввода-вывода перечня сигналов — каналы модулей, обмен Modbus, адаптеры ПЧ. Адресов %I/%Q в
// коде нет: каналы привязываются в дереве устройств (I/O Mapping → «Map to existing variable»), значения Modbus пишет и
// читает слой Modbus, переменные ПЧ — адаптеры приложения (docs/MANUAL_STEPS.md).
{attribute 'qualified_only'}
VAR_GLOBAL
    // === Входы модулей ввода-вывода (DI, AI): дерево устройств, I/O Mapping → Map to existing variable ===
    rLT101_mA : REAL;  // A1.1 · LT101 · Уровень в приёмном резервуаре · 0…5 м
    rPT201_mA : REAL;  // A1.2 · PT201 · Давление в напорном коллекторе · 0…10 бар
    rFT202_mA : REAL;  // A1.3 · FT202 · Расход в напорном коллекторе · 0…500 м³/ч
    rAT401_mA : REAL;  // A1.4 · AT401 · Концентрация сероводорода H₂S в павильоне · 0…40 мг/м³
    rAT402_mA : REAL;  // A1.5 · AT402 · Концентрация метана CH₄ в павильоне · 0…100 % НКПР
    xLS102 : BOOL;  // D1.1 · LS102 · Поплавок «аварийно высокий уровень» (H, 4,2 м)
    xLS103 : BOOL;  // D1.2 · LS103 · Поплавок «сухой ход» (L, 0,4 м)
    xLS203 : BOOL;  // D1.3 · LS203 · Затопление камеры задвижек
    xES301 : BOOL;  // D1.4 · ES301 · Напряжение на вводе в норме (реле контроля фаз)
    xYS302 : BOOL;  // D1.5 · YS302 · ИБП шкафа управления: работа от батарей
    xYS303 : BOOL;  // D1.6 · YS303 · ИБП шкафа управления: неисправность или разряд батарей
    xZS404 : BOOL;  // D1.7 · ZS404 · Дверь павильона открыта
    xYS405 : BOOL;  // D1.8 · YS405 · Пожар (сигнал прибора пожарной сигнализации)
    xHS501 : BOOL;  // D1.9 · HS501 · Кнопка «Сброс аварий» на двери шкафа управления
    xHS502 : BOOL;  // D1.10 · HS502 · Кнопка «Отключить звук» на двери шкафа управления
    xV1_RFB : BOOL;  // D1.11 · V1_RFB · Вентилятор В1: в работе (блок-контакт пускателя)
    xV1_FLT : BOOL;  // D1.12 · V1_FLT · Вентилятор В1: авария (автомат защиты двигателя)
    xP101_RFB : BOOL;  // D2.1 · P101_RFB · Насос Н1: ПЧ в работе (релейный выход ПЧ)
    xP101_FLT : BOOL;  // D2.2 · P101_FLT · Насос Н1: авария ПЧ (релейный выход ПЧ)
    xHS114 : BOOL;  // D2.3 · HS114 · Насос Н1: переключатель «Местное/Дистанционное» в положении «Местное»
    xTS112 : BOOL;  // D2.4 · TS112 · Насос Н1: перегрев обмотки (термовыключатели, реле защиты насоса)
    xMS113 : BOOL;  // D2.5 · MS113 · Насос Н1: протечка в камеру статора (датчик влажности, реле защиты насоса)
    xP102_RFB : BOOL;  // D2.6 · P102_RFB · Насос Н2: ПЧ в работе (релейный выход ПЧ)
    xP102_FLT : BOOL;  // D2.7 · P102_FLT · Насос Н2: авария ПЧ (релейный выход ПЧ)
    xHS124 : BOOL;  // D2.8 · HS124 · Насос Н2: переключатель «Местное/Дистанционное» в положении «Местное»
    xTS122 : BOOL;  // D2.9 · TS122 · Насос Н2: перегрев обмотки (термовыключатели, реле защиты насоса)
    xMS123 : BOOL;  // D2.10 · MS123 · Насос Н2: протечка в камеру статора (датчик влажности, реле защиты насоса)
    xP103_RFB : BOOL;  // D2.11 · P103_RFB · Насос Н3: ПЧ в работе (релейный выход ПЧ)
    xP103_FLT : BOOL;  // D2.12 · P103_FLT · Насос Н3: авария ПЧ (релейный выход ПЧ)
    xHS134 : BOOL;  // D2.13 · HS134 · Насос Н3: переключатель «Местное/Дистанционное» в положении «Местное»
    xTS132 : BOOL;  // D2.14 · TS132 · Насос Н3: перегрев обмотки (термовыключатели, реле защиты насоса)
    xMS133 : BOOL;  // D2.15 · MS133 · Насос Н3: протечка в камеру статора (датчик влажности, реле защиты насоса)

    // === Выходы модулей ввода-вывода (DO, AO): дерево устройств, I/O Mapping → Map to existing variable ===
    xP101_RUN : BOOL;  // Q1.1 · P101_RUN · Насос Н1: команда «Работа» на ПЧ
    xP102_RUN : BOOL;  // Q1.2 · P102_RUN · Насос Н2: команда «Работа» на ПЧ
    xP103_RUN : BOOL;  // Q1.3 · P103_RUN · Насос Н3: команда «Работа» на ПЧ
    xV1_RUN : BOOL;  // Q1.4 · V1_RUN · Вентилятор В1: команда «Работа»
    xHA1 : BOOL;  // Q1.5 · HA1 · Сирена на шкафу управления · без ФБ — код приложения
    xHL1 : BOOL;  // Q1.6 · HL1 · Лампа «Авария» на двери шкафа управления · без ФБ — код приложения
    xK1 : BOOL;  // Q1.7 · K1 · Реле «Общая авария» (сухой контакт в диспетчерскую) · без ФБ — код приложения

    // === Modbus, ПЛК — master, чтение: значения пишет слой Modbus ===
    wP101_STW : WORD;  // RS485-1 · слейв 1 · FC3 4x 100 WORD · P101_STW · Насос Н1: слово состояния ПЧ · адаптер ПЧ
    // RS485-1 · слейв 1 · FC3 4x 101 UINT · P101_FACT · Насос Н1: фактическая частота ПЧ · 0…50 Гц · адаптер ПЧ
    uiP101_FACT : UINT;
    uiIT111 : UINT;  // RS485-1 · слейв 1 · FC3 4x 102 UINT · IT111 · Насос Н1: ток двигателя (измеряет ПЧ) · 0…60 А
    // RS485-1 · слейв 1 · FC3 4x 103 UINT · P101_FCODE · Насос Н1: код последней аварии ПЧ (читает адаптер ПЧ) · без ФБ
    // — код приложения
    uiP101_FCODE : UINT;
    wP102_STW : WORD;  // RS485-1 · слейв 2 · FC3 4x 100 WORD · P102_STW · Насос Н2: слово состояния ПЧ · адаптер ПЧ
    // RS485-1 · слейв 2 · FC3 4x 101 UINT · P102_FACT · Насос Н2: фактическая частота ПЧ · 0…50 Гц · адаптер ПЧ
    uiP102_FACT : UINT;
    uiIT121 : UINT;  // RS485-1 · слейв 2 · FC3 4x 102 UINT · IT121 · Насос Н2: ток двигателя (измеряет ПЧ) · 0…60 А
    // RS485-1 · слейв 2 · FC3 4x 103 UINT · P102_FCODE · Насос Н2: код последней аварии ПЧ (читает адаптер ПЧ) · без ФБ
    // — код приложения
    uiP102_FCODE : UINT;
    wP103_STW : WORD;  // RS485-1 · слейв 3 · FC3 4x 100 WORD · P103_STW · Насос Н3: слово состояния ПЧ · адаптер ПЧ
    // RS485-1 · слейв 3 · FC3 4x 101 UINT · P103_FACT · Насос Н3: фактическая частота ПЧ · 0…50 Гц · адаптер ПЧ
    uiP103_FACT : UINT;
    uiIT131 : UINT;  // RS485-1 · слейв 3 · FC3 4x 102 UINT · IT131 · Насос Н3: ток двигателя (измеряет ПЧ) · 0…60 А
    // RS485-1 · слейв 3 · FC3 4x 103 UINT · P103_FCODE · Насос Н3: код последней аварии ПЧ (читает адаптер ПЧ) · без ФБ
    // — код приложения
    uiP103_FCODE : UINT;
    rTT403 : REAL;  // RS485-2 · слейв 10 · FC4 3x 0 REAL HL · TT403 · Температура воздуха в павильоне · -40…60 °C

    // === Modbus, ПЛК — master, запись: значения читает слой Modbus ===
    wP101_CTW : WORD;  // RS485-1 · слейв 1 · FC16 4x 0 WORD · P101_CTW · Насос Н1: слово управления ПЧ · адаптер ПЧ
    // RS485-1 · слейв 1 · FC16 4x 1 UINT · P101_FREF · Насос Н1: задание частоты ПЧ · 0…50 Гц · адаптер ПЧ
    uiP101_FREF : UINT;
    wP102_CTW : WORD;  // RS485-1 · слейв 2 · FC16 4x 0 WORD · P102_CTW · Насос Н2: слово управления ПЧ · адаптер ПЧ
    // RS485-1 · слейв 2 · FC16 4x 1 UINT · P102_FREF · Насос Н2: задание частоты ПЧ · 0…50 Гц · адаптер ПЧ
    uiP102_FREF : UINT;
    wP103_CTW : WORD;  // RS485-1 · слейв 3 · FC16 4x 0 WORD · P103_CTW · Насос Н3: слово управления ПЧ · адаптер ПЧ
    // RS485-1 · слейв 3 · FC16 4x 1 UINT · P103_FREF · Насос Н3: задание частоты ПЧ · 0…50 Гц · адаптер ПЧ
    uiP103_FREF : UINT;

    // === Состояние обмена со слейвами: пишет слой Modbus (TRUE — обмен исправен) ===
    xMbOk_RS485_1_S1 : BOOL;  // линия RS485-1, слейв 1: обмен исправен
    xMbOk_RS485_1_S2 : BOOL;  // линия RS485-1, слейв 2: обмен исправен
    xMbOk_RS485_1_S3 : BOOL;  // линия RS485-1, слейв 3: обмен исправен
    xMbOk_RS485_2_S10 : BOOL;  // линия RS485-2, слейв 10: обмен исправен

    // === Адаптеры ПЧ (код приложения) → ФБ: разобранное слово состояния и фактическая скорость ===
    xP101_CommOk : BOOL;  // P101: обмен с ПЧ исправен → xCommOk
    xP101_VfdRun : BOOL;  // P101: ПЧ в работе (слово состояния) → xVfdRunning
    xP101_VfdReady : BOOL;  // P101: ПЧ готов к пуску (слово состояния) → xVfdReady
    xP101_VfdFault : BOOL;  // P101: авария ПЧ (слово состояния) → xVfdFault
    rP101_SpeedAct_pct : REAL;  // P101: фактическая скорость, % → rSpeedAct_pct
    xP102_CommOk : BOOL;  // P102: обмен с ПЧ исправен → xCommOk
    xP102_VfdRun : BOOL;  // P102: ПЧ в работе (слово состояния) → xVfdRunning
    xP102_VfdReady : BOOL;  // P102: ПЧ готов к пуску (слово состояния) → xVfdReady
    xP102_VfdFault : BOOL;  // P102: авария ПЧ (слово состояния) → xVfdFault
    rP102_SpeedAct_pct : REAL;  // P102: фактическая скорость, % → rSpeedAct_pct
    xP103_CommOk : BOOL;  // P103: обмен с ПЧ исправен → xCommOk
    xP103_VfdRun : BOOL;  // P103: ПЧ в работе (слово состояния) → xVfdRunning
    xP103_VfdReady : BOOL;  // P103: ПЧ готов к пуску (слово состояния) → xVfdReady
    xP103_VfdFault : BOOL;  // P103: авария ПЧ (слово состояния) → xVfdFault
    rP103_SpeedAct_pct : REAL;  // P103: фактическая скорость, % → rSpeedAct_pct

    // === ФБ → адаптеры ПЧ: задание скорости и команды для слова управления ===
    rP101_SpeedRef_pct : REAL;  // P101: задание на ПЧ, % ← rSpeedRef_pct
    xP101_VfdQRun : BOOL;  // P101: команда «работа» для слова управления ← xQRun
    xP101_VfdQReset : BOOL;  // P101: импульс сброса аварии ПЧ для слова управления ← xQReset
    rP102_SpeedRef_pct : REAL;  // P102: задание на ПЧ, % ← rSpeedRef_pct
    xP102_VfdQRun : BOOL;  // P102: команда «работа» для слова управления ← xQRun
    xP102_VfdQReset : BOOL;  // P102: импульс сброса аварии ПЧ для слова управления ← xQReset
    rP103_SpeedRef_pct : REAL;  // P103: задание на ПЧ, % ← rSpeedRef_pct
    xP103_VfdQRun : BOOL;  // P103: команда «работа» для слова управления ← xQRun
    xP103_VfdQReset : BOOL;  // P103: импульс сброса аварии ПЧ для слова управления ← xQReset
END_VAR

(* ---- GVL_Persist.pvl.st ---- *)
// AUTO-GENERATED by iolistgen 0.2.0 — не редактировать; источник: 03_io_list.csv
// SHA-256 перечня 06336d13c4b2; генератор st-codesys
// Назначение: объект Persistent Variables (контракт plc-process-lib 18.3): Cfg и Retain устройств, по переменной на
// устройство, по возрастанию dev_no. Новое устройство — dev_no больше прежних (переменные встают в конец); типы
// существующих переменных не меняются. Начальные значения — уставки перечня; после загрузки действуют сохранённые
// значения, уставки проекта применяет PRG_ApplyProjectCfg. После устройств — данные приложения (persist_extra), новые —
// в конец. Объект создаётся в CODESYS вручную (docs/MANUAL_STEPS.md); «Reorder List and Clear Gaps» не выполнять.
VAR_GLOBAL PERSISTENT RETAIN
    uiLayoutVersion : UINT := 1;  // версия раскладки списка
    // --- dev_no 11: P101 — Насос Н1 (MotorVfd) ---
    stP101Cfg : PL.ST_MotorCfg := (
        tFbStart := T#10S,
        tFbStop := T#15S,
        tMinStop := T#30S,
        uiMaxStartsPerHour := 10,
        stVfd := (
            rSpeedMin_pct := 60.0,
            rRampUp_pctps := 5.0,
            rRampDown_pctps := 5.0,
            xFbFromComm := FALSE,
            xCommLossIsFault := FALSE
        ),
        udiAlarmIdBase := 110
    );
    stP101Retain : PL.ST_DeviceRetain;  // режим, вывод из работы, наработка, операции
    // --- dev_no 12: P102 — Насос Н2 (MotorVfd) ---
    stP102Cfg : PL.ST_MotorCfg := (
        tFbStart := T#10S,
        tFbStop := T#15S,
        tMinStop := T#30S,
        uiMaxStartsPerHour := 10,
        stVfd := (
            rSpeedMin_pct := 60.0,
            rRampUp_pctps := 5.0,
            rRampDown_pctps := 5.0,
            xFbFromComm := FALSE,
            xCommLossIsFault := FALSE
        ),
        udiAlarmIdBase := 120
    );
    stP102Retain : PL.ST_DeviceRetain;  // режим, вывод из работы, наработка, операции
    // --- dev_no 13: P103 — Насос Н3 (MotorVfd) ---
    stP103Cfg : PL.ST_MotorCfg := (
        tFbStart := T#10S,
        tFbStop := T#15S,
        tMinStop := T#30S,
        uiMaxStartsPerHour := 10,
        stVfd := (
            rSpeedMin_pct := 60.0,
            rRampUp_pctps := 5.0,
            rRampDown_pctps := 5.0,
            xFbFromComm := FALSE,
            xCommLossIsFault := FALSE
        ),
        udiAlarmIdBase := 130
    );
    stP103Retain : PL.ST_DeviceRetain;  // режим, вывод из работы, наработка, операции
    // --- dev_no 14: V1 — Вытяжной вентилятор В1 павильона (Motor) ---
    stV1Cfg : PL.ST_MotorCfg := (
        tMinStop := T#10S,
        udiAlarmIdBase := 140,
        astAlarm := [
            (ePriority := PL.E_AlarmPriority.Low),  // 0 FailToStart
            (ePriority := PL.E_AlarmPriority.Low),  // 1 FeedbackLost
            (ePriority := PL.E_AlarmPriority.High),  // 2 FailToStop
            (ePriority := PL.E_AlarmPriority.High),  // 3 UncommandedRun
            (ePriority := PL.E_AlarmPriority.Low),  // 4 ExtFault
            (ePriority := PL.E_AlarmPriority.None),  // 5 InterlockTrip
            (ePriority := PL.E_AlarmPriority.Medium),  // 6 CommLoss
            (ePriority := PL.E_AlarmPriority.Low)  // 7 SpeedDeviation
        ]
    );
    stV1Retain : PL.ST_DeviceRetain;  // режим, вывод из работы, наработка, операции
    // --- dev_no 101: LT101 — Уровень в приёмном резервуаре (AnalogInput, без Retain) ---
    stLT101Cfg : PL.ST_AnalogInputCfg := (
        rRangeHi_eu := 5.0,
        tFilter := T#2S,
        astLimit := [
            (xEnable := TRUE, rSetpoint_eu := 4.0, rHyst_eu := 0.05, tOnDelay := T#3S),  // 0 HH
            (xEnable := TRUE, rSetpoint_eu := 3.5, rHyst_eu := 0.05, tOnDelay := T#3S),  // 1 H
            (xEnable := TRUE, rSetpoint_eu := 0.8, rHyst_eu := 0.05, tOnDelay := T#3S),  // 2 L
            (xEnable := TRUE, rSetpoint_eu := 0.5, rHyst_eu := 0.05, tOnDelay := T#3S)  // 3 LL
        ],
        udiAlarmIdBase := 1010,
        astAlarm := [
            (ePriority := PL.E_AlarmPriority.High),  // 0 HH
            (ePriority := PL.E_AlarmPriority.Medium),  // 1 H
            (ePriority := PL.E_AlarmPriority.Medium),  // 2 L
            (ePriority := PL.E_AlarmPriority.High),  // 3 LL
            (ePriority := PL.E_AlarmPriority.Medium),  // 4 Failure
            (ePriority := PL.E_AlarmPriority.Low),  // 5 OutOfRange
            (ePriority := PL.E_AlarmPriority.None),  // 6 (резерв)
            (ePriority := PL.E_AlarmPriority.None)  // 7 (резерв)
        ]
    );
    // --- dev_no 102: LS102 — Поплавок «аварийно высокий уровень» (H, 4,2 м) (DigitalInput, без Retain) ---
    stLS102Cfg : PL.ST_DigitalInputCfg := (
        xInvert := TRUE,
        tOnDelay := T#2S,
        udiAlarmIdBase := 1020,
        astAlarm := [
            (ePriority := PL.E_AlarmPriority.High),  // 0 State
            (ePriority := PL.E_AlarmPriority.Medium),  // 1 Failure
            (ePriority := PL.E_AlarmPriority.None),  // 2 (резерв)
            (ePriority := PL.E_AlarmPriority.None),  // 3 (резерв)
            (ePriority := PL.E_AlarmPriority.None),  // 4 (резерв)
            (ePriority := PL.E_AlarmPriority.None),  // 5 (резерв)
            (ePriority := PL.E_AlarmPriority.None),  // 6 (резерв)
            (ePriority := PL.E_AlarmPriority.None)  // 7 (резерв)
        ]
    );
    // --- dev_no 103: LS103 — Поплавок «сухой ход» (L, 0,4 м) (DigitalInput, без Retain) ---
    stLS103Cfg : PL.ST_DigitalInputCfg := (
        xInvert := TRUE,
        tOnDelay := T#1S,
        eFailValue := PL.E_DiFailValue.ForceTrue,
        udiAlarmIdBase := 1030,
        astAlarm := [
            (ePriority := PL.E_AlarmPriority.High),  // 0 State
            (ePriority := PL.E_AlarmPriority.Medium),  // 1 Failure
            (ePriority := PL.E_AlarmPriority.None),  // 2 (резерв)
            (ePriority := PL.E_AlarmPriority.None),  // 3 (резерв)
            (ePriority := PL.E_AlarmPriority.None),  // 4 (резерв)
            (ePriority := PL.E_AlarmPriority.None),  // 5 (резерв)
            (ePriority := PL.E_AlarmPriority.None),  // 6 (резерв)
            (ePriority := PL.E_AlarmPriority.None)  // 7 (резерв)
        ]
    );
    // --- dev_no 111: IT111 — Насос Н1: ток двигателя (измеряет ПЧ) (AnalogInput, без Retain) ---
    stIT111Cfg : PL.ST_AnalogInputCfg := (
        eInput := PL.E_AiInputType.Raw,
        rRangeHi_eu := 60.0,
        rRawHi_cnt := 600.0,
        tFilter := T#1S,
        astLimit := [
            (xEnable := TRUE, rSetpoint_eu := 34.0, tOnDelay := T#10S),  // 0 HH
            (xEnable := TRUE, rSetpoint_eu := 31.0, tOnDelay := T#10S),  // 1 H
            (xEnable := FALSE),  // 2 L
            (xEnable := FALSE)  // 3 LL
        ],
        udiAlarmIdBase := 1110,
        astAlarm := [
            (ePriority := PL.E_AlarmPriority.Medium),  // 0 HH
            (ePriority := PL.E_AlarmPriority.Low),  // 1 H
            (ePriority := PL.E_AlarmPriority.Low),  // 2 L
            (ePriority := PL.E_AlarmPriority.Medium),  // 3 LL
            (ePriority := PL.E_AlarmPriority.Medium),  // 4 Failure
            (ePriority := PL.E_AlarmPriority.Low),  // 5 OutOfRange
            (ePriority := PL.E_AlarmPriority.None),  // 6 (резерв)
            (ePriority := PL.E_AlarmPriority.None)  // 7 (резерв)
        ]
    );
    // --- dev_no 112: TS112 — Насос Н1: перегрев обмотки (термовыключатели, реле защиты… (DigitalInput, без Retain) ---
    stTS112Cfg : PL.ST_DigitalInputCfg := (
        xInvert := TRUE,
        udiAlarmIdBase := 1120,
        astAlarm := [
            (ePriority := PL.E_AlarmPriority.High),  // 0 State
            (ePriority := PL.E_AlarmPriority.Medium),  // 1 Failure
            (ePriority := PL.E_AlarmPriority.None),  // 2 (резерв)
            (ePriority := PL.E_AlarmPriority.None),  // 3 (резерв)
            (ePriority := PL.E_AlarmPriority.None),  // 4 (резерв)
            (ePriority := PL.E_AlarmPriority.None),  // 5 (резерв)
            (ePriority := PL.E_AlarmPriority.None),  // 6 (резерв)
            (ePriority := PL.E_AlarmPriority.None)  // 7 (резерв)
        ]
    );
    // --- dev_no 113: MS113 — Насос Н1: протечка в камеру статора (датчик влажности, ре… (DigitalInput, без Retain) ---
    stMS113Cfg : PL.ST_DigitalInputCfg := (
        tOnDelay := T#10S,
        udiAlarmIdBase := 1130,
        astAlarm := [
            (ePriority := PL.E_AlarmPriority.Medium),  // 0 State
            (ePriority := PL.E_AlarmPriority.Medium),  // 1 Failure
            (ePriority := PL.E_AlarmPriority.None),  // 2 (резерв)
            (ePriority := PL.E_AlarmPriority.None),  // 3 (резерв)
            (ePriority := PL.E_AlarmPriority.None),  // 4 (резерв)
            (ePriority := PL.E_AlarmPriority.None),  // 5 (резерв)
            (ePriority := PL.E_AlarmPriority.None),  // 6 (резерв)
            (ePriority := PL.E_AlarmPriority.None)  // 7 (резерв)
        ]
    );
    // --- dev_no 121: IT121 — Насос Н2: ток двигателя (измеряет ПЧ) (AnalogInput, без Retain) ---
    stIT121Cfg : PL.ST_AnalogInputCfg := (
        eInput := PL.E_AiInputType.Raw,
        rRangeHi_eu := 60.0,
        rRawHi_cnt := 600.0,
        tFilter := T#1S,
        astLimit := [
            (xEnable := TRUE, rSetpoint_eu := 34.0, tOnDelay := T#10S),  // 0 HH
            (xEnable := TRUE, rSetpoint_eu := 31.0, tOnDelay := T#10S),  // 1 H
            (xEnable := FALSE),  // 2 L
            (xEnable := FALSE)  // 3 LL
        ],
        udiAlarmIdBase := 1210,
        astAlarm := [
            (ePriority := PL.E_AlarmPriority.Medium),  // 0 HH
            (ePriority := PL.E_AlarmPriority.Low),  // 1 H
            (ePriority := PL.E_AlarmPriority.Low),  // 2 L
            (ePriority := PL.E_AlarmPriority.Medium),  // 3 LL
            (ePriority := PL.E_AlarmPriority.Medium),  // 4 Failure
            (ePriority := PL.E_AlarmPriority.Low),  // 5 OutOfRange
            (ePriority := PL.E_AlarmPriority.None),  // 6 (резерв)
            (ePriority := PL.E_AlarmPriority.None)  // 7 (резерв)
        ]
    );
    // --- dev_no 122: TS122 — Насос Н2: перегрев обмотки (термовыключатели, реле защиты… (DigitalInput, без Retain) ---
    stTS122Cfg : PL.ST_DigitalInputCfg := (
        xInvert := TRUE,
        udiAlarmIdBase := 1220,
        astAlarm := [
            (ePriority := PL.E_AlarmPriority.High),  // 0 State
            (ePriority := PL.E_AlarmPriority.Medium),  // 1 Failure
            (ePriority := PL.E_AlarmPriority.None),  // 2 (резерв)
            (ePriority := PL.E_AlarmPriority.None),  // 3 (резерв)
            (ePriority := PL.E_AlarmPriority.None),  // 4 (резерв)
            (ePriority := PL.E_AlarmPriority.None),  // 5 (резерв)
            (ePriority := PL.E_AlarmPriority.None),  // 6 (резерв)
            (ePriority := PL.E_AlarmPriority.None)  // 7 (резерв)
        ]
    );
    // --- dev_no 123: MS123 — Насос Н2: протечка в камеру статора (датчик влажности, ре… (DigitalInput, без Retain) ---
    stMS123Cfg : PL.ST_DigitalInputCfg := (
        tOnDelay := T#10S,
        udiAlarmIdBase := 1230,
        astAlarm := [
            (ePriority := PL.E_AlarmPriority.Medium),  // 0 State
            (ePriority := PL.E_AlarmPriority.Medium),  // 1 Failure
            (ePriority := PL.E_AlarmPriority.None),  // 2 (резерв)
            (ePriority := PL.E_AlarmPriority.None),  // 3 (резерв)
            (ePriority := PL.E_AlarmPriority.None),  // 4 (резерв)
            (ePriority := PL.E_AlarmPriority.None),  // 5 (резерв)
            (ePriority := PL.E_AlarmPriority.None),  // 6 (резерв)
            (ePriority := PL.E_AlarmPriority.None)  // 7 (резерв)
        ]
    );
    // --- dev_no 131: IT131 — Насос Н3: ток двигателя (измеряет ПЧ) (AnalogInput, без Retain) ---
    stIT131Cfg : PL.ST_AnalogInputCfg := (
        eInput := PL.E_AiInputType.Raw,
        rRangeHi_eu := 60.0,
        rRawHi_cnt := 600.0,
        tFilter := T#1S,
        astLimit := [
            (xEnable := TRUE, rSetpoint_eu := 34.0, tOnDelay := T#10S),  // 0 HH
            (xEnable := TRUE, rSetpoint_eu := 31.0, tOnDelay := T#10S),  // 1 H
            (xEnable := FALSE),  // 2 L
            (xEnable := FALSE)  // 3 LL
        ],
        udiAlarmIdBase := 1310,
        astAlarm := [
            (ePriority := PL.E_AlarmPriority.Medium),  // 0 HH
            (ePriority := PL.E_AlarmPriority.Low),  // 1 H
            (ePriority := PL.E_AlarmPriority.Low),  // 2 L
            (ePriority := PL.E_AlarmPriority.Medium),  // 3 LL
            (ePriority := PL.E_AlarmPriority.Medium),  // 4 Failure
            (ePriority := PL.E_AlarmPriority.Low),  // 5 OutOfRange
            (ePriority := PL.E_AlarmPriority.None),  // 6 (резерв)
            (ePriority := PL.E_AlarmPriority.None)  // 7 (резерв)
        ]
    );
    // --- dev_no 132: TS132 — Насос Н3: перегрев обмотки (термовыключатели, реле защиты… (DigitalInput, без Retain) ---
    stTS132Cfg : PL.ST_DigitalInputCfg := (
        xInvert := TRUE,
        udiAlarmIdBase := 1320,
        astAlarm := [
            (ePriority := PL.E_AlarmPriority.High),  // 0 State
            (ePriority := PL.E_AlarmPriority.Medium),  // 1 Failure
            (ePriority := PL.E_AlarmPriority.None),  // 2 (резерв)
            (ePriority := PL.E_AlarmPriority.None),  // 3 (резерв)
            (ePriority := PL.E_AlarmPriority.None),  // 4 (резерв)
            (ePriority := PL.E_AlarmPriority.None),  // 5 (резерв)
            (ePriority := PL.E_AlarmPriority.None),  // 6 (резерв)
            (ePriority := PL.E_AlarmPriority.None)  // 7 (резерв)
        ]
    );
    // --- dev_no 133: MS133 — Насос Н3: протечка в камеру статора (датчик влажности, ре… (DigitalInput, без Retain) ---
    stMS133Cfg : PL.ST_DigitalInputCfg := (
        tOnDelay := T#10S,
        udiAlarmIdBase := 1330,
        astAlarm := [
            (ePriority := PL.E_AlarmPriority.Medium),  // 0 State
            (ePriority := PL.E_AlarmPriority.Medium),  // 1 Failure
            (ePriority := PL.E_AlarmPriority.None),  // 2 (резерв)
            (ePriority := PL.E_AlarmPriority.None),  // 3 (резерв)
            (ePriority := PL.E_AlarmPriority.None),  // 4 (резерв)
            (ePriority := PL.E_AlarmPriority.None),  // 5 (резерв)
            (ePriority := PL.E_AlarmPriority.None),  // 6 (резерв)
            (ePriority := PL.E_AlarmPriority.None)  // 7 (резерв)
        ]
    );
    // --- dev_no 201: PT201 — Давление в напорном коллекторе (AnalogInput, без Retain) ---
    stPT201Cfg : PL.ST_AnalogInputCfg := (
        rRangeHi_eu := 10.0,
        tFilter := T#1S,
        astLimit := [
            (xEnable := TRUE, rSetpoint_eu := 5.0, tOnDelay := T#5S),  // 0 HH
            (xEnable := TRUE, rSetpoint_eu := 4.0, tOnDelay := T#5S),  // 1 H
            (xEnable := TRUE, rSetpoint_eu := 1.0, rHyst_eu := 0.1, tOnDelay := T#5S),  // 2 L
            (xEnable := TRUE, rSetpoint_eu := 0.5, rHyst_eu := 0.1, tOnDelay := T#5S)  // 3 LL
        ],
        udiAlarmIdBase := 2010,
        astAlarm := [
            (ePriority := PL.E_AlarmPriority.High),  // 0 HH
            (ePriority := PL.E_AlarmPriority.Medium),  // 1 H
            (ePriority := PL.E_AlarmPriority.Medium),  // 2 L
            (ePriority := PL.E_AlarmPriority.High),  // 3 LL
            (ePriority := PL.E_AlarmPriority.Medium),  // 4 Failure
            (ePriority := PL.E_AlarmPriority.Low),  // 5 OutOfRange
            (ePriority := PL.E_AlarmPriority.None),  // 6 (резерв)
            (ePriority := PL.E_AlarmPriority.None)  // 7 (резерв)
        ]
    );
    // --- dev_no 202: FT202 — Расход в напорном коллекторе (AnalogInput, без Retain) ---
    stFT202Cfg : PL.ST_AnalogInputCfg := (
        rRangeHi_eu := 500.0,
        rLowCut_pct := 1.0,
        tFilter := T#3S,
        astLimit := [
            (xEnable := FALSE),  // 0 HH
            (xEnable := FALSE),  // 1 H
            (xEnable := TRUE, rSetpoint_eu := 30.0, rHyst_eu := 5.0, tOnDelay := T#30S),  // 2 L
            (xEnable := FALSE)  // 3 LL
        ],
        udiAlarmIdBase := 2020,
        astAlarm := [
            (ePriority := PL.E_AlarmPriority.High),  // 0 HH
            (ePriority := PL.E_AlarmPriority.Low),  // 1 H
            (ePriority := PL.E_AlarmPriority.Medium),  // 2 L
            (ePriority := PL.E_AlarmPriority.High),  // 3 LL
            (ePriority := PL.E_AlarmPriority.Medium),  // 4 Failure
            (ePriority := PL.E_AlarmPriority.Low),  // 5 OutOfRange
            (ePriority := PL.E_AlarmPriority.None),  // 6 (резерв)
            (ePriority := PL.E_AlarmPriority.None)  // 7 (резерв)
        ]
    );
    // --- dev_no 203: LS203 — Затопление камеры задвижек (DigitalInput, без Retain) ---
    stLS203Cfg : PL.ST_DigitalInputCfg := (
        tOnDelay := T#5S,
        udiAlarmIdBase := 2030,
        astAlarm := [
            (ePriority := PL.E_AlarmPriority.Medium),  // 0 State
            (ePriority := PL.E_AlarmPriority.Medium),  // 1 Failure
            (ePriority := PL.E_AlarmPriority.None),  // 2 (резерв)
            (ePriority := PL.E_AlarmPriority.None),  // 3 (резерв)
            (ePriority := PL.E_AlarmPriority.None),  // 4 (резерв)
            (ePriority := PL.E_AlarmPriority.None),  // 5 (резерв)
            (ePriority := PL.E_AlarmPriority.None),  // 6 (резерв)
            (ePriority := PL.E_AlarmPriority.None)  // 7 (резерв)
        ]
    );
    // --- dev_no 301: ES301 — Напряжение на вводе в норме (реле контроля фаз) (DigitalInput, без Retain) ---
    stES301Cfg : PL.ST_DigitalInputCfg := (
        tOnDelay := T#3S,
        xAlarmOnTrue := FALSE,
        udiAlarmIdBase := 3010,
        astAlarm := [
            (ePriority := PL.E_AlarmPriority.High),  // 0 State
            (ePriority := PL.E_AlarmPriority.Medium),  // 1 Failure
            (ePriority := PL.E_AlarmPriority.None),  // 2 (резерв)
            (ePriority := PL.E_AlarmPriority.None),  // 3 (резерв)
            (ePriority := PL.E_AlarmPriority.None),  // 4 (резерв)
            (ePriority := PL.E_AlarmPriority.None),  // 5 (резерв)
            (ePriority := PL.E_AlarmPriority.None),  // 6 (резерв)
            (ePriority := PL.E_AlarmPriority.None)  // 7 (резерв)
        ]
    );
    // --- dev_no 302: YS302 — ИБП шкафа управления: работа от батарей (DigitalInput, без Retain) ---
    stYS302Cfg : PL.ST_DigitalInputCfg := (
        tOnDelay := T#5S,
        udiAlarmIdBase := 3020,
        astAlarm := [
            (ePriority := PL.E_AlarmPriority.Medium),  // 0 State
            (ePriority := PL.E_AlarmPriority.Medium),  // 1 Failure
            (ePriority := PL.E_AlarmPriority.None),  // 2 (резерв)
            (ePriority := PL.E_AlarmPriority.None),  // 3 (резерв)
            (ePriority := PL.E_AlarmPriority.None),  // 4 (резерв)
            (ePriority := PL.E_AlarmPriority.None),  // 5 (резерв)
            (ePriority := PL.E_AlarmPriority.None),  // 6 (резерв)
            (ePriority := PL.E_AlarmPriority.None)  // 7 (резерв)
        ]
    );
    // --- dev_no 303: YS303 — ИБП шкафа управления: неисправность или разряд батарей (DigitalInput, без Retain) ---
    stYS303Cfg : PL.ST_DigitalInputCfg := (
        tOnDelay := T#5S,
        udiAlarmIdBase := 3030,
        astAlarm := [
            (ePriority := PL.E_AlarmPriority.Medium),  // 0 State
            (ePriority := PL.E_AlarmPriority.Medium),  // 1 Failure
            (ePriority := PL.E_AlarmPriority.None),  // 2 (резерв)
            (ePriority := PL.E_AlarmPriority.None),  // 3 (резерв)
            (ePriority := PL.E_AlarmPriority.None),  // 4 (резерв)
            (ePriority := PL.E_AlarmPriority.None),  // 5 (резерв)
            (ePriority := PL.E_AlarmPriority.None),  // 6 (резерв)
            (ePriority := PL.E_AlarmPriority.None)  // 7 (резерв)
        ]
    );
    // --- dev_no 401: AT401 — Концентрация сероводорода H₂S в павильоне (AnalogInput, без Retain) ---
    stAT401Cfg : PL.ST_AnalogInputCfg := (
        rRangeHi_eu := 40.0,
        astLimit := [
            (xEnable := TRUE, rSetpoint_eu := 10.0, rHyst_eu := 0.5, tOnDelay := T#5S),  // 0 HH
            (xEnable := TRUE, rSetpoint_eu := 5.0, rHyst_eu := 0.5, tOnDelay := T#5S),  // 1 H
            (xEnable := FALSE),  // 2 L
            (xEnable := FALSE)  // 3 LL
        ],
        udiAlarmIdBase := 4010,
        astAlarm := [
            (ePriority := PL.E_AlarmPriority.High),  // 0 HH
            (ePriority := PL.E_AlarmPriority.Medium),  // 1 H
            (ePriority := PL.E_AlarmPriority.Medium),  // 2 L
            (ePriority := PL.E_AlarmPriority.High),  // 3 LL
            (ePriority := PL.E_AlarmPriority.Medium),  // 4 Failure
            (ePriority := PL.E_AlarmPriority.Low),  // 5 OutOfRange
            (ePriority := PL.E_AlarmPriority.None),  // 6 (резерв)
            (ePriority := PL.E_AlarmPriority.None)  // 7 (резерв)
        ]
    );
    // --- dev_no 402: AT402 — Концентрация метана CH₄ в павильоне (AnalogInput, без Retain) ---
    stAT402Cfg : PL.ST_AnalogInputCfg := (
        astLimit := [
            (xEnable := TRUE, rSetpoint_eu := 20.0, rHyst_eu := 1.0, tOnDelay := T#5S),  // 0 HH
            (xEnable := TRUE, rSetpoint_eu := 10.0, rHyst_eu := 1.0, tOnDelay := T#5S),  // 1 H
            (xEnable := FALSE),  // 2 L
            (xEnable := FALSE)  // 3 LL
        ],
        udiAlarmIdBase := 4020,
        astAlarm := [
            (ePriority := PL.E_AlarmPriority.High),  // 0 HH
            (ePriority := PL.E_AlarmPriority.Medium),  // 1 H
            (ePriority := PL.E_AlarmPriority.Medium),  // 2 L
            (ePriority := PL.E_AlarmPriority.High),  // 3 LL
            (ePriority := PL.E_AlarmPriority.Medium),  // 4 Failure
            (ePriority := PL.E_AlarmPriority.Low),  // 5 OutOfRange
            (ePriority := PL.E_AlarmPriority.None),  // 6 (резерв)
            (ePriority := PL.E_AlarmPriority.None)  // 7 (резерв)
        ]
    );
    // --- dev_no 403: TT403 — Температура воздуха в павильоне (AnalogInput, без Retain) ---
    stTT403Cfg : PL.ST_AnalogInputCfg := (
        eInput := PL.E_AiInputType.Eng,
        rRangeLo_eu := -40.0,
        rRangeHi_eu := 60.0,
        astLimit := [
            (xEnable := FALSE),  // 0 HH
            (xEnable := TRUE, rSetpoint_eu := 35.0, rHyst_eu := 1.0, tOnDelay := T#1M),  // 1 H
            (xEnable := TRUE, rSetpoint_eu := 5.0, rHyst_eu := 1.0, tOnDelay := T#1M),  // 2 L
            (xEnable := FALSE)  // 3 LL
        ],
        udiAlarmIdBase := 4030,
        astAlarm := [
            (ePriority := PL.E_AlarmPriority.Low),  // 0 HH
            (ePriority := PL.E_AlarmPriority.Low),  // 1 H
            (ePriority := PL.E_AlarmPriority.Low),  // 2 L
            (ePriority := PL.E_AlarmPriority.Low),  // 3 LL
            (ePriority := PL.E_AlarmPriority.Medium),  // 4 Failure
            (ePriority := PL.E_AlarmPriority.Low),  // 5 OutOfRange
            (ePriority := PL.E_AlarmPriority.None),  // 6 (резерв)
            (ePriority := PL.E_AlarmPriority.None)  // 7 (резерв)
        ]
    );
    // --- dev_no 404: ZS404 — Дверь павильона открыта (DigitalInput, без Retain) ---
    stZS404Cfg : PL.ST_DigitalInputCfg := (
        tOnDelay := T#2S,
        udiAlarmIdBase := 4040,
        astAlarm := [
            (ePriority := PL.E_AlarmPriority.Low),  // 0 State
            (ePriority := PL.E_AlarmPriority.Medium),  // 1 Failure
            (ePriority := PL.E_AlarmPriority.None),  // 2 (резерв)
            (ePriority := PL.E_AlarmPriority.None),  // 3 (резерв)
            (ePriority := PL.E_AlarmPriority.None),  // 4 (резерв)
            (ePriority := PL.E_AlarmPriority.None),  // 5 (резерв)
            (ePriority := PL.E_AlarmPriority.None),  // 6 (резерв)
            (ePriority := PL.E_AlarmPriority.None)  // 7 (резерв)
        ]
    );
    // --- dev_no 405: YS405 — Пожар (сигнал прибора пожарной сигнализации) (DigitalInput, без Retain) ---
    stYS405Cfg : PL.ST_DigitalInputCfg := (
        udiAlarmIdBase := 4050,
        astAlarm := [
            (ePriority := PL.E_AlarmPriority.High),  // 0 State
            (ePriority := PL.E_AlarmPriority.Medium),  // 1 Failure
            (ePriority := PL.E_AlarmPriority.None),  // 2 (резерв)
            (ePriority := PL.E_AlarmPriority.None),  // 3 (резерв)
            (ePriority := PL.E_AlarmPriority.None),  // 4 (резерв)
            (ePriority := PL.E_AlarmPriority.None),  // 5 (резерв)
            (ePriority := PL.E_AlarmPriority.None),  // 6 (резерв)
            (ePriority := PL.E_AlarmPriority.None)  // 7 (резерв)
        ]
    );
    // --- dev_no 501: HS501 — Кнопка «Сброс аварий» на двери шкафа управления (DigitalInput, без Retain) ---
    stHS501Cfg : PL.ST_DigitalInputCfg := (udiAlarmIdBase := 5010);
    // --- dev_no 502: HS502 — Кнопка «Отключить звук» на двери шкафа управления (DigitalInput, без Retain) ---
    stHS502Cfg : PL.ST_DigitalInputCfg := (udiAlarmIdBase := 5020);
    // --- данные приложения, persist_extra (persist_station.txt): новые — только в конец ---
    stStationCfg : ST_StationCfg;  // уставки станции (04 §18.2, № 2–31)
    stStationRetain : ST_StationRetain;  // режим, способ, следующий ведущий
    // LIC101 (04 §18.2, № 32–43)
    stLIC101Cfg : PL.ST_PidCfg := (eAction := PL.E_PidAction.Direct, rKp := 6.0, rTi_s := 600.0, rTd_s := 0.0, rPvMin_eu := 0.0, rPvMax_eu := 5.0, rSpMin_eu := 1.2, rSpMax_eu := 2.2, rOutMin_pct := 0.0, rOutMax_pct := 100.0, tSample := T#500MS, ePvFailAction := PL.E_PidPvFailAction.Hold, rSafeOut_pct := 100.0, xUseOutAct := TRUE, udiAlarmIdBase := 100100, astAlarm := [(ePriority := PL.E_AlarmPriority.None), (ePriority := PL.E_AlarmPriority.None), (ePriority := PL.E_AlarmPriority.None), (ePriority := PL.E_AlarmPriority.None), (ePriority := PL.E_AlarmPriority.None), (ePriority := PL.E_AlarmPriority.None), (ePriority := PL.E_AlarmPriority.None), (ePriority := PL.E_AlarmPriority.None)]);
    stLIC101Retain : PL.ST_DeviceRetain;  // режим регулятора
    stStationCfgLkg : ST_StationCfg;  // последняя корректная копия уставок станции (LKG): переживает перезапуск
END_VAR
